Fanuc KAREL source: kx00027.KL

-- PROVISIONAL review KL for V770-1; original PC SHA256 7726a4890fb6d59c49cca0890d77302df2eadaa8c80f2ac19ded18b3c4eb7d53
-- Incomplete behavior may be omitted. Consult companion uncertainty JSON. Do not deploy.
PROGRAM KX00027
%NOLOCKGROUP
VAR
  I : INTEGER
  J : INTEGER
  B : BOOLEAN
  F : FILE
  S : STRING[80]
-- UNRESOLVED_DECL P type=000102
BEGIN
  -- UNRESOLVED_PC offsets 5-12; opcodes 9D,23
  -- UNRESOLVED_PC offsets 17-21; opcodes 7F
END KX00027
